(* IEC 61131-3 sources: stc/examples, 3 files *)

(* ---- comments.st ---- *)
PROGRAM comments
// single line comment
  VAR // end of line comment
  END_VAR (* comment *)

(* start comment
this is a multiline comment
end comment *)

END_PROGRAM;

(* ---- empty_program.st ---- *)
PROGRAM emptyprogram
  VAR
  END_VAR

END_PROGRAM;

(* ---- variable_declaration.st ---- *)
PROGRAM variabledeclaration
  VAR
    x : BOOL;
  END_VAR
  x := TRUE;
END_PROGRAM;
